{attribute 'qualified_only'}
VAR_GLOBAL
	gHoming : ST_HomingResult;
END_VAR

(* stored: Version 1.1.0.1, ProductVersion 3.1.4024.15
   GVL GVL_HomingResult: Id {12bbacfe-0286-4811-80b5-4a925471803a} *)
